Fanuc KAREL source: KA00068.KL

PROGRAM KA00068
%NOLOCKGROUP
VAR
  SRC: XYZWPR
  DST: JOINTPOS
BEGIN
  SRC.X = 1.0
  DST = SRC
END KA00068
